  rq_init_comm_if_connected(9, "1")
  rq_init_comm_if_connected(2, "2")
  rq_init_comm_if_connected(3, "3")
  rq_init_comm_if_connected(4, "4")
  rq_print_connected_grippers()
  rq_gripper_communication_thread = run rq_gripper_communication()
  set_closed_norm(97.6470588235294, 1)
  set_open_norm(1.1764705882352942, 1)
  set_closed_mm(0.0, 1)
  set_open_mm(53.0, 1)
  set_closed_norm(100.0, 2)
  set_open_norm(0.0, 2)
  set_closed_mm(0.0, 2)
  set_open_mm(50.0, 2)
  set_closed_norm(100.0, 3)
  set_open_norm(0.0, 3)
  set_closed_mm(0.0, 3)
  set_open_mm(50.0, 3)
  set_closed_norm(100.0, 4)
  set_open_norm(0.0, 4)
  set_closed_mm(0.0, 4)
  set_open_mm(50.0, 4)
  rq_current_limit_enabled = False
  while(not rq_gripper_communication_thread_started):
      sync()
  end
  # end: URCap Installation Node
  step_count_adf59958_3206_4157_9784_b10371ce5c7f = 0.0
  thread Step_Counter_Thread_24389c08_1df7_4ce5_b554_c14c432d27df():
    while (True):
      step_count_adf59958_3206_4157_9784_b10371ce5c7f = step_count_adf59958_3206_4157_9784_b10371ce5c7f + 1.0
      sync()
    end
  end
  run Step_Counter_Thread_24389c08_1df7_4ce5_b554_c14c432d27df()
  global easyPickCount_1=0
  global easyPickCount_2=0
  global easyPickNoObj_1=0
  global easyPickNoObj_2=0
  global easyPickParts_1=0
  global easyPickParts_2=0
  global Waypoint_5_p=p[-.503981135492, -.020518307034, -.008276831947, .000014057113, -.000040888691, -1.552034036819]
  global Waypoint_5_q=[-2.833382291967979, -1.9212651814221733, -2.1321875237240953, -0.6588229253369251, 1.5722038270431158, -2.850154288451896]
  global Waypoint_6_p=p[-.503981135427, -.020518307013, .254365481595, .000014057113, -.000040888692, -1.552034036819]
  global Waypoint_6_q=[-2.8325741195847134, -1.5732649512396772, -1.7571224084645864, -1.3818883320232143, 1.5731996450940247, -2.8512813934633954]
  while (True):
    $ 2 "Robot Program"
    $ 3 "Home (Safe)"
    movej([-1.2302089344500047, -1.2969853503591224, -1.875639182904262, -1.539621866126728, 1.5731943360401213, -2.80099559440227], a=1.3962634015954636, v=1.0471975511965976)
    # begin: URCap Program Node
    #   Source: SensoPart VISOR Robotic, 2.0.0, SensoPart Industriesensorik GmbH
    #   Type: VISOR Robotic App
    $ 38 "VISOR Easy Pick"
    def visorFuncEasyPick_d89785():
      # begin: URCap Program Node
      #   Source: SensoPart VISOR Robotic, 2.0.0, SensoPart Industriesensorik GmbH
      #   Type: Easy Pick Setup
      $ 39 "# 1 Setup" "noBreak"
      local easyPickVisorId = 1
      local easyPickArmMounted = True
      local easyPickSetJob = True
      local easyPickJobName = "Spatula_1"
      local easyPickAtImgAcq = False
      local easyPickImgAcqPose = p[-0.6152,-0.0058,0.3709,0.0000,0.0000,-1.6045]
      # end: URCap Program Node
      # begin: URCap Program Node
      #   Source: SensoPart VISOR Robotic, 2.0.0, SensoPart Industriesensorik GmbH
      #   Type: Process
      $ 40 "Process" "noBreak"
      local easyPickObjTaken = False
      local easyPickTrigger = False
      local easyPickPoseIdx = 0
      local easyPickPose = p[0,0,0,0,0,0]
      def easyPickFuncTrigger(visorId, setJob, jobName, arm):
      if (setJob):
        visor_changeJob(visorId, jobName, 6000)
      end
      if (arm):
        visor_trigger(visorId, 6000, "arm")
      else:
        visor_trigger(visorId, 6000)
      end
      global easyPickParts_2=visor_partsFound(visorId)
      visor_easyPickUpdate(visorId, "parts", visor_partsFound(visorId))
      return visor_getPose3d(visorId, 0)
    end
    while (not easyPickObjTaken):
      easyPickTrigger = (easyPickCount_2 >= visor_partsFound(easyPickVisorId)) or (easyPickCount_2 > 9) or (not visor_easyPickCheckIdent("0a25a2", easyPickVisorId))
      if (easyPickTrigger):
        easyPickCount_2 = 0
      end
      easyPickPoseIdx = easyPickCount_2
      easyPickPose = visor_getPose3d(easyPickVisorId, easyPickPoseIdx)
      visor_easyPickUpdate(easyPickVisorId, "counter", easyPickPoseIdx)
      # begin: URCap Program Node
      #   Source: SensoPart VISOR Robotic, 2.0.0, SensoPart Industriesensorik GmbH
      #   Type: Image Acquisition Pose
      $ 41 "Image Acquisition Pose" "noBreak"
      if (easyPickTrigger):
        if (not easyPickAtImgAcq):
          movej(pose_trans(easyPickImgAcqPose,p[0.0000,0.0000,-0.0000,0.0000,0.0000,0.0000]),a=1.3963,v=1.0472,t=0.000000,r=0.000000)
          easyPickAtImgAcq = True
        end
        easyPickPose = easyPickFuncTrigger(easyPickVisorId, easyPickSetJob, easyPickJobName, easyPickArmMounted)
      end
      # end: URCap Program Node
      # begin: URCap Program Node
      #   Source: SensoPart VISOR Robotic, 2.0.0, SensoPart Industriesensorik GmbH
      #   Type: Object Detected
      $ 42 "Object Detected" "noBreak"
      if (visor_partsFound(easyPickVisorId) > 0):
        $ 43 "Open Gripper" "noBreak"
        # begin: URCap Program Node
        #   Source: Robotiq_Grippers, 1.8.4.4844, Robotiq Inc.
        #   Type: Gripper
        $ 44 "Gripper Move40mm (1)" "noBreak"
        if not(gripper_connected[0]):
          popup("Gripper 1 must be connected to run this program.", "No connection", False, True, True)
        end
        if not(rq_is_gripper_activated("1")):
          popup("Gripper 1 is not activated. Go to Installation tab > Gripper to activate it and run the program again.", "Not activated", False, True, True)
        end
        rq_set_pos_spd_for(63, 92, 77, "1")
        rq_wait_pos_spe_for_request(63, 92, 77, "1")
        rq_go_to("1")
        rq_wait("1")
        # end: URCap Program Node
        # begin: URCap Program Node
        #   Source: SensoPart VISOR Robotic, 2.0.0, SensoPart Industriesensorik GmbH
        #   Type: Approach Pose
        $ 45 "Approach Pose" "noBreak"
        movej(pose_trans(easyPickPose,p[0.0000,0.0000,0.0700,0.0000,0.0000,0.0000]),a=1.3963,v=1.0472,t=0.000000,r=0.000000)
        # end: URCap Program Node
        # begin: URCap Program Node
        #   Source: SensoPart VISOR Robotic, 2.0.0, SensoPart Industriesensorik GmbH
        #   Type: Target Pose
        $ 46 "Target Pose" "noBreak"
        movel(pose_trans(easyPickPose,p[0.0000,0.0000,-0.0000,0.0000,0.0000,0.0000]),a=0.5000,v=0.2500,t=0.000000,r=0.000000)
        # end: URCap Program Node
        $ 47 "Close Gripper" "noBreak"
        # begin: URCap Program Node
        #   Source: Robotiq_Grippers, 1.8.4.4844, Robotiq Inc.
        #   Type: Gripper
        $ 48 "Gripper Close (1)" "noBreak"
        if not(gripper_connected[0]):
          popup("Gripper 1 must be connected to run this program.", "No connection", False, True, True)
        end
        if not(rq_is_gripper_activated("1")):
          popup("Gripper 1 is not activated. Go to Installation tab > Gripper to activate it and run the program again.", "Not activated", False, True, True)
        end
        rq_set_pos_spd_for(255, 92, 77, "1")
        rq_wait_pos_spe_for_request(255, 92, 77, "1")
        rq_go_to("1")
        rq_wait("1")
        # end: URCap Program Node
        # begin: URCap Program Node
        #   Source: SensoPart VISOR Robotic, 2.0.0, SensoPart Industriesensorik GmbH
        #   Type: Exit Pose
        $ 49 "Exit Pose" "noBreak"
        movel(pose_trans(easyPickPose,p[0.0000,0.0000,-0.0000,0.0000,0.0000,0.0000]),a=0.5000,v=0.2500,t=0.000000,r=0.000000)
        # end: URCap Program Node
        easyPickObjTaken = True
      end
      # end: URCap Program Node
      # begin: URCap Program Node
      #   Source: SensoPart VISOR Robotic, 2.0.0, SensoPart Industriesensorik GmbH
      #   Type: No Object Detected
      $ 50 "No Object Detected" "noBreak"
      if (visor_partsFound(easyPickVisorId) < 1):
        $ 51 "Popup: No object detected" "noBreak"
        popup("No object detected", "Message", False, False, blocking=True)
        else:
      end
      # end: URCap Program Node
    end
    easyPickCount_2 = easyPickCount_2 + 1
    visor_easyPickUpdate(easyPickVisorId, "counter", easyPickCount_2)
    visor_easyPickSetIdent("0a25a2", easyPickVisorId)
    # end: URCap Program Node
  end
  visorFuncEasyPick_d89785()
  # end: URCap Program Node
  $ 52 "MoveJ"
  $ 53 "Waypoint_5" "breakAfter"
  movej(get_inverse_kin(Waypoint_5_p, qnear=Waypoint_5_q), a=1.3962634015954636, v=1.0471975511965976)
  $ 54 "Waypoint_6" "breakAfter"
  movej(get_inverse_kin(Waypoint_6_p, qnear=Waypoint_6_q), a=1.3962634015954636, v=1.0471975511965976)
  $ 55 "Home (Safe)"
  movej([-1.2302089344500047, -1.2969853503591224, -1.875639182904262, -1.539621866126728, 1.5731943360401213, -2.80099559440227], a=1.3962634015954636, v=1.0471975511965976)
  # begin: URCap Program Node
  #   Source: Robotiq_Grippers, 1.8.4.4844, Robotiq Inc.
  #   Type: Gripper
  $ 56 "Gripper Open (1)"
  if not(gripper_connected[0]):
    popup("Gripper 1 must be connected to run this program.", "No connection", False, True, True)
  end
  if not(rq_is_gripper_activated("1")):
    popup("Gripper 1 is not activated. Go to Installation tab > Gripper to activate it and run the program again.", "Not activated", False, True, True)
  end
  rq_set_pos_spd_for(0, 92, 77, "1")
  rq_wait_pos_spe_for_request(0, 92, 77, "1")
  rq_go_to("1")
  rq_wait("1")
  # end: URCap Program Node
  end
end
